(* IEC 61131-3 sources: kns-port-domestic/tools/inventory_tests/fixtures/app/src/POUs/PRG_Example, 1 file *)

(* ---- PRG_Example.decl.st ---- *)
// Назначение: пример шаблона
PROGRAM PRG_Example
VAR
    xRun : BOOL;
END_VAR
